(* IEC 61131-3 sources: plcassist-cli/packages/volt-lsp-iec/test-corpus/pro2193/Device/Plc Logic/Application/09 Misc/Library Manager/L_MC2P_MotionControlCam (part 2) *)

(* ---- L_MC2P_TEMPLATEAXIS.fb ---- *)
FUNCTION_BLOCK L_MC2P_TEMPLATEAXIS
VAR_IN_OUT
	AXIS : AXIS_REF;
END_VAR
VAR
	SINSTANCESTR : STRING;
	XERROROLD : BOOL;
	WERRORIDOLD : WORD;
	DWERRORITFID : DWORD;
END_VAR
END_FUNCTION_BLOCK

METHOD FB_GETERRORITFID : DWORD
END_METHOD

METHOD FB_RESETERROR
VAR_INPUT
	XERROR : BOOL;
	WERRORID : WORD;
END_VAR
END_METHOD

METHOD FB_SETERROR
VAR_INPUT
	WERRORID : WORD := 0;
	XSETERRORSTOP : BOOL := FALSE;
END_VAR
END_METHOD

METHOD FB_INIT : BOOL
VAR_INPUT
	BINITRETAINS : BOOL;
	BINCOPYCODE : BOOL;
END_VAR
END_METHOD

(* ---- L_MC2P_TEMPLATEAXIS_LICENCE.fb ---- *)
FUNCTION_BLOCK L_MC2P_TEMPLATEAXIS_LICENCE EXTENDS L_MC2P_TemplateAxis
VAR
	LICHANDLING : L_IMHP_LLMHandling;
END_VAR
END_FUNCTION_BLOCK

METHOD ACTIVATEAPPCREDIT : BOOL
VAR_INPUT
	XACTIVATE : BOOL;
END_VAR
END_METHOD

(* ---- L_MC2P_TEMPLATEMASTERAXIS.fb ---- *)
FUNCTION_BLOCK L_MC2P_TEMPLATEMASTERAXIS
VAR_IN_OUT
	MASTER : AXIS_REF;
END_VAR
VAR
	SINSTANCESTR : STRING;
	XERROROLD : BOOL;
	WERRORIDOLD : WORD;
	DWERRORITFID : DWORD;
END_VAR
END_FUNCTION_BLOCK

METHOD FB_GETERRORITFID : DWORD
END_METHOD

METHOD FB_RESETERROR
VAR_INPUT
	XERROR : BOOL;
	WERRORID : WORD;
END_VAR
END_METHOD

METHOD FB_SETERROR
VAR_INPUT
	WERRORID : WORD := 0;
	XSETERRORSTOP : BOOL := FALSE;
END_VAR
END_METHOD

METHOD FB_INIT : BOOL
VAR_INPUT
	BINITRETAINS : BOOL;
	BINCOPYCODE : BOOL;
END_VAR
END_METHOD

(* ---- L_MC2P_TEMPLATENOAXIS.fb ---- *)
FUNCTION_BLOCK L_MC2P_TEMPLATENOAXIS
VAR
	SINSTANCESTR : STRING;
	XERROROLD : BOOL;
	WERRORIDOLD : WORD;
END_VAR
END_FUNCTION_BLOCK

METHOD FB_INIT : BOOL
VAR_INPUT
	BINITRETAINS : BOOL;
	BINCOPYCODE : BOOL;
END_VAR
END_METHOD

(* ---- L_MC2P_TEMPLATESLAVEAXIS.fb ---- *)
FUNCTION_BLOCK L_MC2P_TEMPLATESLAVEAXIS
VAR_IN_OUT
	SLAVE : AXIS_REF;
END_VAR
VAR
	SINSTANCESTR : STRING;
	XERROROLD : BOOL;
	WERRORIDOLD : WORD;
	DWERRORITFID : DWORD;
END_VAR
END_FUNCTION_BLOCK

METHOD FB_GETERRORITFID : DWORD
END_METHOD

METHOD FB_RESETERROR
VAR_INPUT
	XERROR : BOOL;
	WERRORID : WORD;
END_VAR
END_METHOD

METHOD FB_SETERROR
VAR_INPUT
	WERRORID : WORD := 0;
	XSETERRORSTOP : BOOL := FALSE;
END_VAR
END_METHOD

METHOD FB_INIT : BOOL
VAR_INPUT
	BINITRETAINS : BOOL;
	BINCOPYCODE : BOOL;
END_VAR
END_METHOD

(* ---- L_MC2P_WRITELMDFILE.fb ---- *)
FUNCTION_BLOCK L_MC2P_WRITELMDFILE
VAR
	TEST1 : BOOL;
	TEST2 : BOOL;
	TEST3 : BOOL;
	TEST4 : BOOL;
	SFILE_INT : STRING := '';
	EDATA_INT : L_MC2P_LMData;
	PDATA_INT : POINTER TO BYTE;
	WDATAELEMENTS_INT : WORD;
	XENABLEONLINECHANGE_INT : BOOL;
	XBUSY_INT : BOOL;
	XDONE_INT : BOOL;
	XERROR_INT : BOOL;
	EERRORID_INT : L_IE1P_Error;
	XEXECUTEOLD : BOOL;
	HFILE : SYSFILE.RTS_IEC_HANDLE;
	RES : SYSFILE.RTS_IEC_RESULT;
	ID : L_MC2P_Magic;
	DWLENGTH : DWORD;
	XACTIVECRYPTING : BOOL;
	CRYPT : Crypting;
	CK : ARRAY [0..3] OF ULINT;
	CCYCLES : WORD;
	DICDATAWRITE : DINT;
	DWSTARTCDATA : DWORD;
	ABDATA : ARRAY [0..15] OF BYTE;
	DATAIDX : DWORD;
	AVAILABLEDATA : DWORD;
	XDATAWRITEDONE : BOOL;
	UDIFSIZE : UDINT;
	UDIFBYTESWRITE : UDINT;
	RELOAD : BOOL;
END_VAR
END_FUNCTION_BLOCK

METHOD CLOSECRYPTFRAME
VAR_INPUT
	HFILE : SYSFILE.RTS_IEC_HANDLE;
END_VAR
END_METHOD

METHOD MAIN
END_METHOD

METHOD OPENCRYPTFRAME
VAR_INPUT
	HFILE : SYSFILE.RTS_IEC_HANDLE;
END_VAR
END_METHOD

METHOD RESET
END_METHOD

METHOD SETDATALENGTH
VAR_INPUT
	HFILE : SYSFILE.RTS_IEC_HANDLE;
END_VAR
END_METHOD

METHOD WRITEFRAMES
VAR_INPUT
	HFILE : SYSFILE.RTS_IEC_HANDLE;
END_VAR
END_METHOD

METHOD WRITEORGA
VAR_INPUT
	HFILE : SYSFILE.RTS_IEC_HANDLE;
END_VAR
END_METHOD

METHOD WRITESPECIFICDATA
VAR_INPUT
	HFILE : SYSFILE.RTS_IEC_HANDLE;
END_VAR
END_METHOD

METHOD CALCCRC : DWORD
VAR_INPUT
	HFILE : SYSFILE.RTS_IEC_HANDLE;
	DWLENGTH : DWORD;
END_VAR
END_METHOD

METHOD CRCCHECKSUM32BITINCREMENTAL : DWORD
VAR_INPUT
	PBDATA : POINTER TO BYTE;
	DWDATASIZE : DWORD;
	DWCRC : DWORD;
END_VAR
END_METHOD

METHOD RESETWRITEDATA
END_METHOD

METHOD CWRITECHAR
VAR_INPUT
	HFILE : SYSFILE.RTS_IEC_HANDLE;
	SDATA : STRING(16);
	N : UINT;
END_VAR
END_METHOD

METHOD CWRITEF64
VAR_INPUT
	HFILE : SYSFILE.RTS_IEC_HANDLE;
	LRDATA : LREAL;
END_VAR
END_METHOD

METHOD CWRITEU16
VAR_INPUT
	HFILE : SYSFILE.RTS_IEC_HANDLE;
	WDATA : WORD;
END_VAR
END_METHOD

METHOD CWRITEU32
VAR_INPUT
	HFILE : SYSFILE.RTS_IEC_HANDLE;
	DWDATA : DWORD;
END_VAR
END_METHOD

METHOD WRITECRYPTDATA : DWORD
VAR_INPUT
	HFILE : SYSFILE.RTS_IEC_HANDLE;
	DWSIZE : DWORD;
END_VAR
VAR_IN_OUT
	DATA : L_MC2P_IntData;
END_VAR
END_METHOD

METHOD WRITE
VAR_INPUT
	HFILE : SYSFILE.RTS_IEC_HANDLE;
	PBYBUFFER : POINTER TO BYTE;
	ULSIZE : UINT;
END_VAR
VAR_OUTPUT
	UDIDATAWRITE : UDINT;
END_VAR
END_METHOD

METHOD WRITECHAR : STRING(16)
VAR_INPUT
	HFILE : SYSFILE.RTS_IEC_HANDLE;
	SDATA : STRING(16);
	N : UINT;
END_VAR
END_METHOD

METHOD WRITEF64 : LREAL
VAR_INPUT
	HFILE : SYSFILE.RTS_IEC_HANDLE;
	LRDATA : LREAL;
END_VAR
END_METHOD

METHOD WRITEU16 : WORD
VAR_INPUT
	HFILE : SYSFILE.RTS_IEC_HANDLE;
	WDATA : WORD;
END_VAR
END_METHOD

METHOD WRITEU32
VAR_INPUT
	HFILE : SYSFILE.RTS_IEC_HANDLE;
	DWDATA : DWORD;
END_VAR
END_METHOD

METHOD ABORT : UDINT
END_METHOD

METHOD EXECUTE : UDINT
END_METHOD

(* ---- MC_CAMIN.fb ---- *)
FUNCTION_BLOCK MC_CAMIN EXTENDS L_MC2P_MasterSlaveSync
VAR_INPUT
	EXECUTE : BOOL;
	CONTINUOUSUPDATE : BOOL := FALSE;
	MASTEROFFSET : LREAL := 0;
	SLAVEOFFSET : LREAL := 0;
	MASTERSCALING : LREAL := 1;
	SLAVESCALING : LREAL := 1;
	MASTERSTARTDISTANCE : LREAL;
	MASTERSYNCPOSITION : LREAL;
	STARTMODE : MC_START_MODE := MC_Start_Mode.mcAbsolute;
	MASTERVALUESOURCE : MC_SOURCE := MC_SOURCE.mcSetValue;
	CAMTABLE : MC_CAM_REF;
	BUFFERMODE : MC_BUFFER_MODE := MC_Buffer_Mode.mcAborting;
	DIRECTCHANGE : BOOL := FALSE;
	CLUTCHTIME : LREAL := 0.001;
	VELOCITYDIFF : LREAL := 3600.0;
	ACCELERATION : LREAL := 3600.0;
	DECELERATION : LREAL := 3600.0;
	JERK : LREAL := 0.0;
	SCALINGOFFSETMODE : L_MC2P_ScalingOffsetMode := L_MC2P_ScalingOffsetMode.direct;
	PERIODIC : BOOL := TRUE;
	MASTERABSOLUTE : BOOL := TRUE;
	SLAVEABSOLUTE : BOOL := TRUE;
END_VAR
VAR_OUTPUT
	INSYNC : BOOL;
	BUSY : BOOL;
	ACTIVE : BOOL;
	COMMANDABORTED : BOOL;
	ERROR : BOOL;
	ERRORID : L_IE1P_Error;
	ENDOFPROFILE : BOOL;
END_VAR
VAR
	XPERIODIC_INT : BOOL;
	XMASTERABSOLUTE_INT : BOOL;
	XSLAVEABSOLUTE_INT : BOOL;
	PSCCAMDATA : POINTER TO L_MC2P_CamData;
	L_MC2P_FLEXCAMSTATE1 : L_MC2P_FlexCamState;
	SCINPUTMASTERSOURCE : L_MC2P_AxisProfile;
	SCACTSLAVE : L_MC2P_AxisProfile;
	SCOUTPUTSLAVE : L_MC2P_AxisProfile;
	EOFFSETMODE_INT : L_MC2P_OffsetMode;
	ESCALINGMODE_INT : L_MC2P_ScalingMode;
	ECLUTCHMODE_INT : L_MC2P_ClutchMode;
	EPOSCTRLDIRECTION_INT : L_MC2P_ReverseCtrlDirection;
	LRMASTEROFFSET_INT : LREAL;
	LRSLAVEOFFSET_INT : LREAL;
	LRMASTERSCALING_INT : LREAL;
	LRSLAVESCALING_INT : LREAL;
	LRMASTERSTARTDISTANCE_INT : LREAL;
	LRMASTERSYNCPOSITION_INT : LREAL;
	ESTARTMODE_INT : MC_START_MODE;
	EMASTERVALUESOURCE_INT : MC_SOURCE;
	EMASTERVALUESOURCE_OLD : MC_SOURCE;
	SCCAMTABLE_INT : MC_CAM_REF;
	SCCAMINFO_INT : L_MC2P_CamInfo;
	ESCALINGOFFSETMODE_INT : L_MC2P_ScalingOffsetMode;
	LRVELOCITYDIFF_INT : LREAL;
	LRACCELERATION_INT : LREAL;
	LRDECELERATION_INT : LREAL;
	LRJERK_INT : LREAL;
	XDIRECTCHANGE_INT : BOOL := FALSE;
	LRCLUTCHTIME_INT : LREAL;
	DWCHANGEID : DWORD := 1;
	STARTINCURRENTPERIOD : BOOL;
END_VAR
END_FUNCTION_BLOCK

METHOD CONVERT_CLOSEMODE
END_METHOD

METHOD CONVERT_SCALINGOFFSETMODE
END_METHOD

METHOD GET_MASTERVALUES
END_METHOD

METHOD READINPUTS
VAR_INPUT
	XREADALL : BOOL;
END_VAR
VAR_IN_OUT
	AXIS : AXIS_REF;
END_VAR
END_METHOD

METHOD RESET_OUTPUTSADD
END_METHOD

METHOD RESET_OUTPUTSBYCOMMANDABORTED
END_METHOD

METHOD RESET_OUTPUTSBYERROR
END_METHOD

METHOD SYNCIN
END_METHOD

METHOD FB_INIT : BOOL
VAR_INPUT
	BINITRETAINS : BOOL;
	BINCOPYCODE : BOOL;
END_VAR
END_METHOD

(* ---- MC_CAMOUT.fb ---- *)
FUNCTION_BLOCK MC_CAMOUT EXTENDS L_MC2P_TemplateSlaveAxis
VAR_INPUT
	EXECUTE : BOOL;
END_VAR
VAR_OUTPUT
	DONE : BOOL;
	BUSY : BOOL;
	ERROR : BOOL;
	ERRORID : L_IE1P_Error;
END_VAR
VAR
	L_MC2P_CLUTCHBASIC1 : L_MC2P_ClutchBasic;
	XSUPERIMPOSED : BOOL;
	WFUNID : WORD;
	SCINPUTSLAVE : L_MC2P_AxisProfile;
	SCOUTPUTSLAVE : L_MC2P_AxisProfile;
	XEXECUTEOLD : BOOL;
	XRESETOUTPUT : BOOL;
	LRJERK : LREAL;
	XDONEINTERN : BOOL;
	XDONEFLAG : BOOL;
END_VAR
END_FUNCTION_BLOCK

METHOD GET_SLAVEJERK
END_METHOD

METHOD GET_SLAVEVALUES
END_METHOD

METHOD RESET_OUTPUTS
END_METHOD

METHOD RESET_OUTPUTSBYCOMMANDABORTED
END_METHOD

METHOD RESET_OUTPUTSBYERROR
END_METHOD

METHOD SET_SLAVEVALUES
END_METHOD

(* ---- MC_COMBINEAXES.fb ---- *)
FUNCTION_BLOCK MC_COMBINEAXES EXTENDS L_MC2P_Template3Axes_Licence
VAR_INPUT
	EXECUTE : BOOL;
	CONTINUOUSUPDATE : BOOL := FALSE;
	COMBINEMODE : MC_COMBINE_MODE := MC_COMBINE_MODE.mcAddAxes;
	GEARRATIONUMERATORM1 : INT := 1;
	GEARRATIODENOMINATORM1 : UINT := 1;
	GEARRATIONUMERATORM2 : INT := 1;
	GEARRATIODENOMINATORM2 : UINT := 1;
	MASTERVALUESOURCEM1 : MC_SOURCE := MC_SOURCE.mcSetValue;
	MASTERVALUESOURCEM2 : MC_SOURCE := MC_SOURCE.mcSetValue;
	BUFFERMODE : MC_BUFFER_MODE := MC_Buffer_Mode.mcAborting;
	VELOCITY : LREAL := 3600.0;
	ACCELERATION : LREAL := 3600.0;
	DECELERATION : LREAL := 3600.0;
	JERK : LREAL := 0.0;
END_VAR
VAR_OUTPUT
	INSYNC : BOOL;
	BUSY : BOOL;
	ACTIVE : BOOL;
	COMMANDABORTED : BOOL;
	ERROR : BOOL;
	ERRORID : L_IE1P_Error;
END_VAR
VAR
	L_MC2P_CLUTCHBASIC1 : L_MC2P_ClutchBasic;
	L_MC2P_CAMAXISCONVERTER1 : L_MC2P_CamAxisConverter;
	L_MC2P_CAMAXISCONVERTER2 : L_MC2P_CamAxisConverter;
	L_MC2P_CAMAXISCONVERTER3 : L_MC2P_CamAxisConverter;
	L_MC2P_MODIFYAXIS1 : L_MC2P_ModifyAxis;
	L_MC2P_MODIFYAXIS2 : L_MC2P_ModifyAxis;
	XSUPERIMPOSED : BOOL;
	WFUNID : WORD;
	SCINPUTMASTERSOURCE1 : L_MC2P_AxisProfile;
	SCINPUTMASTERSOURCE2 : L_MC2P_AxisProfile;
	SCACTSLAVE : L_MC2P_AxisProfile;
	SCOUTPUTSLAVE : L_MC2P_AxisProfile;
	LRSETSCALING1 : LREAL;
	LRSETSCALING2 : LREAL;
	XEXECUTEOLD : BOOL;
	XCOMMANDABORTEDOLD : BOOL;
	INSYNCOLD : BOOL;
	XRESETOUTPUT : BOOL;
	XCONTINUOUSUPDATE : BOOL;
	XUPDATEBLOCKER : BOOL;
	UIUPDATECOUNTER : UINT;
	XCLUTCHACTIVE : BOOL;
	DWINSTANCE : __XWORD;
	XBUFFERACTIVE : BOOL;
	XPREVBUFFBDONE : BOOL;
	LRPOSOLDMASTER1 : LREAL;
	LRPOSOLDMASTER2 : LREAL;
	LRPOSMODTOLIMMASTER1 : LREAL;
	LRPOSMODTOLIMMASTER2 : LREAL;
	ECOMBINEMODE_INT : MC_COMBINE_MODE;
	IGEARRATIONUMERATORM1_INT : INT;
	UIGEARRATIODENOMINATORM1_INT : UINT := 1;
	IGEARRATIONUMERATORM2_INT : INT;
	UIGEARRATIODENOMINATORM2_INT : UINT := 1;
	EMASTERVALUESOURCEM1_INT : MC_SOURCE;
	EMASTERVALUESOURCEM2_INT : MC_SOURCE;
	LRVELOCITY_INT : LREAL;
	LRACCELERATION_INT : LREAL;
	LRDECELERATION_INT : LREAL;
	LRJERK_INT : LREAL;
	EBUFFERMODE_INT : MC_BUFFER_MODE;
	XERROR_TMP1 : BOOL;
	XERROR_TMP2 : BOOL;
	XERROR_TMP3 : BOOL;
	EERRORID_TMP1 : L_IE1P_Error;
	EERRORID_TMP2 : L_IE1P_Error;
	EERRORID_TMP3 : L_IE1P_Error;
END_VAR
END_FUNCTION_BLOCK

METHOD CALC_COMBINEAXES
END_METHOD

METHOD CHECK_AXISDATA
END_METHOD

METHOD CHECK_CONTINUOUSUPDATE
END_METHOD

METHOD CHECK_FORUPDATES
END_METHOD

METHOD GET_MASTERVALUES
END_METHOD

METHOD GET_SLAVEVALUES
END_METHOD

METHOD LOAD_AXISCONVERTER
END_METHOD

METHOD POSMASTER1MODTOLIM : LREAL
END_METHOD

METHOD POSMASTER2MODTOLIM : LREAL
END_METHOD

METHOD READINPUTS
VAR_INPUT
	XREADALL : BOOL;
END_VAR
END_METHOD

METHOD RESET_OUTPUTS
END_METHOD

METHOD RESET_OUTPUTSBYCOMMANDABORTED
END_METHOD

METHOD RESET_OUTPUTSBYERROR
END_METHOD

METHOD SET_BUFFERMODE
END_METHOD

METHOD SET_SLAVEVALUES
END_METHOD

(* ---- MC_GEARIN.fb ---- *)
FUNCTION_BLOCK MC_GEARIN EXTENDS L_MC2P_MasterSlaveSync
VAR_INPUT
	EXECUTE : BOOL;
	CONTINUOUSUPDATE : BOOL := FALSE;
	RATIONUMERATOR : INT := 1;
	RATIODENOMINATOR : UINT := 1;
	MASTERVALUESOURCE : MC_SOURCE := MC_SOURCE.mcSetValue;
	ACCELERATION : LREAL := 3600.0;
	DECELERATION : LREAL := 3600.0;
	JERK : LREAL := 0.0;
	BUFFERMODE : MC_BUFFER_MODE := MC_Buffer_Mode.mcAborting;
END_VAR
VAR_OUTPUT
	INGEAR : BOOL;
	BUSY : BOOL;
	ACTIVE : BOOL;
	COMMANDABORTED : BOOL;
	ERROR : BOOL;
	ERRORID : L_IE1P_Error;
END_VAR
VAR
	L_MC2P_CLUTCHBASIC1 : L_MC2P_ClutchBasic;
	L_MC2P_MODIFYAXIS1 : L_MC2P_ModifyAxis;
	L_MC2P_AXISCONVERTER1 : L_MC2P_AxisConverterBase;
	SCINPUTMASTERSOURCE : L_MC2P_AxisProfile;
	SCINPUTMASTERSCALED : L_MC2P_AxisProfile;
	SCACTSLAVE : L_MC2P_AxisProfile;
	SCOUTPUTSLAVE : L_MC2P_AxisProfile;
	LRPOSDIFF : LREAL;
	LRSETSCALING : LREAL;
	IRATIONUMERATOR_INT : INT;
	UIRATIODENOMINATOR_INT : UINT := 1;
	EMASTERVALUESOURCE_INT : MC_SOURCE;
	LRACCELERATION_INT : LREAL;
	LRDECELERATION_INT : LREAL;
	LRJERK_INT : LREAL;
	LROFFSET : LREAL;
	_L_MC2P_MASTERCONVERTERTOSLAVELEGTH : L_MC2P_AxisConverterBase;
	_SCINPUTMASTERCONVERTERTED : L_MC2P_AxisProfile;
	_XAXISCONVERTERCONVERTERTED : BOOL;
END_VAR
END_FUNCTION_BLOCK

METHOD CALC_SLAVEVALUES
END_METHOD

METHOD GET_MASTERVALUES
END_METHOD

METHOD READINPUTS
VAR_INPUT
	XREADALL : BOOL;
END_VAR
VAR_IN_OUT
	AXIS : AXIS_REF;
END_VAR
END_METHOD

METHOD RESET_OUTPUTSADD
END_METHOD

METHOD SET_BUFFERMODE
END_METHOD

METHOD SYNCIN
END_METHOD

METHOD FB_INIT : BOOL
VAR_INPUT
	BINITRETAINS : BOOL;
	BINCOPYCODE : BOOL;
END_VAR
END_METHOD

(* ---- MC_GEARINPOS.fb ---- *)
FUNCTION_BLOCK MC_GEARINPOS EXTENDS L_MC2P_MasterSlaveSync
VAR_INPUT
	EXECUTE : BOOL;
	RATIONUMERATOR : INT := 1;
	RATIODENOMINATOR : UINT := 1;
	MASTERVALUESOURCE : MC_SOURCE := MC_SOURCE.mcSetValue;
	MASTERSYNCPOSITION : LREAL;
	SLAVESYNCPOSITION : LREAL;
	SYNCMODE : MC_SYNC_MODE;
	MASTERSTARTDISTANCE : LREAL;
	BUFFERMODE : MC_BUFFER_MODE := MC_Buffer_Mode.mcAborting;
END_VAR
VAR_OUTPUT
	STARTSYNC : BOOL;
	INSYNC : BOOL;
	BUSY : BOOL;
	ACTIVE : BOOL;
	COMMANDABORTED : BOOL;
	ERROR : BOOL;
	ERRORID : L_IE1P_Error;
END_VAR
VAR
	L_MC2P_CLUTCHBASIC1 : L_MC2P_ClutchBasic;
	L_MC2P_MODIFYAXIS1 : L_MC2P_ModifyAxis;
	L_MC2P_AXISCONVERTER1 : L_MC2P_AxisConverterBase;
	SCINPUTMASTERSOURCE : L_MC2P_AxisProfile;
	SCINPUTMASTERSCALED : L_MC2P_AxisProfile;
	SCACTSLAVE : L_MC2P_AxisProfile;
	SCENDSLAVE : L_MC2P_AxisProfile;
	SCOUTPUTSLAVE : L_MC2P_AxisProfile;
	LRPOSDIFF : LREAL;
	LRSETSCALING : LREAL;
	LRCORRECTSYNCMODEPOS : LREAL;
	LRCALCMASTERDISTANCE : LREAL;
	IRATIONUMERATOR_INT : INT;
	UIRATIODENOMINATOR_INT : UINT := 1;
	EMASTERVALUESOURCE_INT : MC_SOURCE;
	LRMASTERSYNCPOSITION_INT : LREAL;
	LRSLAVESYNCPOSITION_INT : LREAL;
	ESYNCMODE_INT : MC_SYNC_MODE;
	LRMASTERSTARTDISTANCE_INT : LREAL;
	LRVELOCITY_INT : LREAL;
	LRACCELERATION_INT : LREAL;
	LRDECELERATION_INT : LREAL;
	LRJERK_INT : LREAL;
	LROFFSET : LREAL;
	DEBUG_INPUTMASTERPOS : LREAL;
	DEBUG_LRMASTERCLUTCHPOSITION : LREAL;
	DEBUG_LRMASTERCLUTCHDISTANCE : LREAL;
	XUSEAXISDIRECTIONINT : BOOL;
	XUSEAXISDIRECTION : BOOL := TRUE;
	USEAXISDIRECTION : BOOL;
END_VAR
END_FUNCTION_BLOCK

METHOD CALC_SLAVEENDVALUES
END_METHOD

METHOD CALC_SLAVEVALUES
END_METHOD

METHOD GET_MASTERVALUES
END_METHOD

METHOD READINPUTS
VAR_INPUT
	XREADALL : BOOL;
END_VAR
VAR_IN_OUT
	AXIS : AXIS_REF;
END_VAR
END_METHOD

METHOD RESET_OUTPUTSADD
END_METHOD

METHOD SET_BUFFERMODE_TEST
END_METHOD

METHOD SYNCIN
END_METHOD

METHOD FB_INIT : BOOL
VAR_INPUT
	BINITRETAINS : BOOL;
	BINCOPYCODE : BOOL;
END_VAR
END_METHOD

(* ---- MC_GEAROUT.fb ---- *)
FUNCTION_BLOCK MC_GEAROUT EXTENDS L_MC2P_TemplateSlaveAxis
VAR_INPUT
	EXECUTE : BOOL;
END_VAR
VAR_OUTPUT
	DONE : BOOL;
	BUSY : BOOL;
	ERROR : BOOL;
	ERRORID : L_IE1P_Error;
END_VAR
VAR
	MC_CAMOUT1 : MC_CamOut;
END_VAR
END_FUNCTION_BLOCK

(* ---- MC_PHASINGABSOLUTE.fb ---- *)
FUNCTION_BLOCK MC_PHASINGABSOLUTE EXTENDS L_MC2P_Phasing
VAR_OUTPUT
	ABSOLUTEPHASESHIFT : LREAL;
END_VAR
END_FUNCTION_BLOCK

(* ---- MC_PHASINGRELATIVE.fb ---- *)
FUNCTION_BLOCK MC_PHASINGRELATIVE EXTENDS L_MC2P_Phasing
VAR_OUTPUT
	COVEREDPHASESHIFT : LREAL;
END_VAR
END_FUNCTION_BLOCK
